(* IEC 61131-3 sources: krc-sample-programs/robot-cell-ethernetip-codesys/source/03_States, 2 files *)

(* ---- E_Step.st ---- *)
// The steps, a thousand apart for the states, a hundred apart for the steps inside a state.
TYPE E_Step :
(
	S0_IDLE           :=    0,	// Idle: powered up and at rest. Goes straight to Not Ready
	S1_NOT_READY      := 1000,	// Not Ready: waiting for the link, the robot, an empty fixture, Stop not pressed
	S2_RESET          := 2000,	// Reset: clears a fault or a stop, waits for Reset to be released
	S3_READY          := 3000,	// Ready: waiting for Start
	S3_STARTING       := 3100,	// Ready: Start pressed, the robot program is starting (play)
	S4_LOAD_REQUEST   := 4000,	// Load: command 1 out, waiting for the robot to acknowledge
	S4_LOADING        := 4100,	// Load: the robot is putting a part in the fixture
	S4_LOAD_CLEAR     := 4200,	// Load: command back to 0, waiting for the robot to clear its answer
	S5_CLAMPING       := 5000,	// Clamping: valve on, setpoint out, waiting for pressure
	S5_HOLDING        := 5100,	// Clamping: at pressure, holding for the hold time
	S6_OPENING        := 6000,	// Opening: valve off, waiting for the clamp to read open
	S7_UNLOAD_REQUEST := 7000,	// Unload: command 2 out, waiting for the robot to acknowledge
	S7_UNLOADING      := 7100,	// Unload: the robot is taking the part out
	S7_UNLOAD_CLEAR   := 7200,	// Unload: command back to 0, waiting for the robot to clear its answer
	S8_FAULT          := 8000,	// Fault: waiting for Reset
	S8_STOPPED        := 8100,	// Stopped: Stop pressed, the robot program stopped (stop), waiting for Reset
	S9_PAUSED         := 9000,	// Paused: Pause pressed, the robot program paused (pause), waiting for Start
	S9_RESUMING       := 9100 	// Paused: Start pressed, the robot program resuming (play)
) INT;
END_TYPE

(* ---- CONSTANTS.st ---- *)
// Named numbers the program uses, so no bare number appears in the logic.
VAR_GLOBAL CONSTANT
	AI_FULL_SCALE    : REAL := 32760.0;	// CC100 analog input raw count at 10 V (WAGO manual, section 9.4)
	AO_FULL_SCALE    : REAL := 32767.0;	// CC100 analog output raw count for 10 V (WAGO manual, section 9.4)
	PRESSURE_RANGE   : REAL := 100.0;	// psi at 10 V, for the sensor and the regulator
	PRESSURE_BAND    : REAL := 2.0;	// psi: within this much of the setpoint counts as at pressure

	// The link: where each word sits in the GVL_Link arrays (the robot's register in the comment).
	TO_HEARTBEAT     : INT := 0;	// Input register 0: PLC heartbeat
	TO_COMMAND       : INT := 1;	// Input register 1: command
	TO_FIXTURE_CLEAR : INT := 2;	// Input register 2: fixture clear
	TO_PLC_STEP      : INT := 3;	// Input register 3: PLC step, for the pendant
	FROM_HEARTBEAT   : INT := 0;	// Output register 0: robot heartbeat
	FROM_READY       : INT := 1;	// Output register 1: robot ready
	FROM_ACK         : INT := 2;	// Output register 2: acknowledge, the command the robot accepted
	FROM_DONE        : INT := 3;	// Output register 3: done, the command the robot finished
	FROM_FAULT       : INT := 4;	// Output register 4: robot fault code
	FROM_ROBOT_STEP  : INT := 5;	// Output register 5: robot step, what the robot program is doing or waiting on
	BIT_START        : INT := 0;	// Input bit register 0: Start (I/O action on the robot)
	BIT_STOP         : INT := 1;	// Input bit register 1: Stop (I/O action on the robot)
	BIT_PAUSE        : INT := 2;	// Input bit register 2: Pause (I/O action on the robot)

	CMD_NONE         : DINT := 0;	// Command: nothing
	CMD_LOAD         : DINT := 1;	// Command: put a part in the fixture
	CMD_UNLOAD       : DINT := 2;	// Command: take the part out
	ROBOT_RUNNING    : SINT := 7;	// Robot mode 7: arm powered, brakes released
	ROBOT_NOT_HOME   : DINT := 900;	// Robot step 900: the program was started away from home and refused to move
	HEARTBEAT_TIME   : TIME := T#250MS;	// How often the PLC counts its heartbeat
	HEARTBEAT_LOST   : TIME := T#1S;	// No change in the robot's heartbeat this long: it's gone
	ROBOT_START_TIME : TIME := T#10S;	// How long the robot program may take to start or resume and be ready
	ROBOT_HOME_CHECK : TIME := T#2S;	// Long enough after Start for the robot program to have written its first step
	ROBOT_PAUSE_TIME : TIME := T#3S;	// How long the robot program may take to pause

	// The Dashboard: the robot's command port.
	ROBOT_IP         : STRING(15) := '192.168.1.10';	// The robot's address (Q2 in the program design), also set in UR_Robot
	DASH_PORT        : UINT := 29999;	// UR's Dashboard Server port
	DASH_POLL_TIME   : TIME := T#250MS;	// How often the PLC asks the robot a question
	DASH_REPLY_TIME  : TIME := T#2S;	// No answer this long: drop the connection and connect again
END_VAR
